// TIA Portal V20 export
// export: Created 2026-10-12T05:14:44.6307195Z, ExportSetting WithDefaults, DisplayName Totally Integrated Automation Portal, DisplayVersion V20, DisplayName TIA Portal Openness, DisplayVersion V20, DisplayName TIA Portal Teamcenter Gateway, DisplayVersion V20, DisplayName TIA Portal Version Control Interface, DisplayVersion V20, DisplayName SINAMICS Startdrive Advanced, DisplayVersion V20 SP1 Update 2, DisplayName SINAMICS Startdrive G110M, G120, G120C, G120D, G120P, G115D, DisplayVersion V20 SP1 Update 2, DisplayName SINAMICS Startdrive G130, G150, S120, S150, SINAMICS MV, G220, S200, S210, DisplayVersion V20 SP1 Update 2, DisplayName STEP 7 Professional, DisplayVersion V20, DisplayName STEP 7 Safety, DisplayVersion V20, DisplayName WinCC Basic/Comfort/Advanced, DisplayVersion V20, DisplayName WinCC Professional, DisplayVersion V20, DisplayName WinCC Unified, DisplayVersion V20
FUNCTION "FRK_UnitMailbox" : Void   // FC72, SCL
{ S7_Optimized_Access := 'TRUE' }
VERSION : 0.1
// stored: AutoNumber true, IsIECCheckEnabled false, SetENOAutomatically false, UDAEnableTagReadback false
   VAR_INPUT
      Supported : Array[0..6] of Bool;
   END_VAR
   VAR_IN_OUT
      Core : "FRK_Core";
      Unit : "FRK_Unit";
      Status : "ST_ModuleStatus";
      Policy : Array[0..6] of "ST_ModePolicy";
      Access : "FRK_Access";
      Request : "ST_HmiRequest";
      Response : "ST_HmiResponse";
   END_VAR
   VAR_TEMP
      SequenceBefore : UDInt;
   END_VAR
BEGIN

   #SequenceBefore := #Request.Sequence;
   IF #SequenceBefore = 0 OR #SequenceBefore = #Unit.SeenSequence THEN
       RETURN;
   END_IF;
   #Unit.Request := #Request;
   IF #Request.Sequence <> #SequenceBefore THEN
       #Unit.Request.Secret := '';
       RETURN;
   END_IF;
   #Request.Secret := '';
   #Unit.RequestUser := #Access.CurrentUser;
   #Unit.SeenSequence := #SequenceBefore;
   #Unit.RequestPending := TRUE;
END_FUNCTION
